// Write side of the event arguments (fluent).
INTERFACE I_ArgumentBuilder

METHOD Clear : I_ArgumentBuilder
END_METHOD

METHOD AddString : I_ArgumentBuilder
VAR_INPUT
	sValue	: T_MaxString;
END_VAR
END_METHOD

METHOD AddDInt : I_ArgumentBuilder
VAR_INPUT
	nValue	: DINT;
END_VAR
END_METHOD

METHOD AddLReal : I_ArgumentBuilder
VAR_INPUT
	fValue		: LREAL;
	nDecimals	: USINT;	// 0..9
END_VAR
END_METHOD

METHOD AddBool : I_ArgumentBuilder
VAR_INPUT
	bValue	: BOOL;
END_VAR
END_METHOD

END_INTERFACE

(* stored: Version 1.1.0.1, ProductVersion 3.1.4026.26
   Itf I_ArgumentBuilder: Id {d52b9beb-7686-498a-a88a-3417ce4241a2}
   Method Clear: Id {848a4de6-37d9-4af5-b1a2-bd4db72c0174}
   Method AddString: Id {7c0d1f56-2379-44ec-a329-b22872f15186}
   Method AddDInt: Id {f77aedb4-6505-4ac4-bd30-df492b671162}
   Method AddLReal: Id {56cc5461-1c86-41e5-85ed-5397c50dbbae}
   Method AddBool: Id {8a1ef3ea-8ff8-4869-9086-92a82127a31c} *)
